FUNCTION FC_FindMax : BOOL

;

END_FUNCTION

(* stored: Version 1.1.0.1, ProductVersion 3.1.4024.12
   POU FC_FindMax: Id {0d5e3531-9289-4021-901d-72888c86c107}, SpecialFunc None *)
